# EPICS substitutions: db/Beckhoff_7XXX/ecmcEX72XX_OPT_csv.substitutions
file "ecmcEL72XX_DRV.template"
{
  pattern {CH_ID, ESLO, EGU}
          {"$(OPT_CH_ID=01)", "$(OPT_VEL_ESLO=2.3406E-5)", "$(OPT_VEL_EGU=rad/s)"}
}
